Staubli VAL3: valGI.pjx

--- valGI.pjx ---
Parameters version=s8.15.3Cs9_BS3337 stackSize=200000 millimeterUnit=true
Program file=_getForce.pgx
Program file=_productCycle.pgx
Program file=_tCycleCtrl.pgx
Program file=createUserTask.pgx
Program file=cycle_Abort.pgx
Program file=cycle_End.pgx
Program file=cycle_GoHome.pgx
Program file=cycle_Hold.pgx
Program file=cycle_Init.pgx
Program file=cycle_Reset.pgx
Program file=cycle_RotGoHome.pgx
Program file=cycle_Start.pgx
Program file=cycle_Stop.pgx
Program file=cycle_Unhold.pgx
Program file=Init.pgx
Program file=kill.pgx
Program file=Main.pgx
Program file=MonitorIO.pgx
Program file=MonitorIO1.pgx
Program file=start.pgx
Program file=stop.pgx
Data file=valGI.dtx
Library alias=rs path=Disk://source/projectSource/robotStatus/robotStatus.pjx
Library alias=io path=Disk://source/projectSource/io/io.pjx
Library alias=act path=Disk://source/projectSource/Action/Action.pjx
Library alias=savedata path=Disk://source/saveData/saveData.pjx
Library alias=home path=Disk://HMI_cs9/home/home.pjx
Library alias=plc path=Disk://source/projectSource/plc/plc.pjx
Library alias=prog path=Disk://source/projectSource/program/program.pjx
Library alias=safeHome path=Disk://source/projectSource/goSafeHome/goSafeHome.pjx
Library alias=safe path=Disk://safeLogic/safeLogic.pjx
Library alias=program path=Disk://source/projectSource/program/program.pjx
Library alias=hmi_util path=Disk://HMI_cs9/HMI_util/HMI_util.pjx
Library alias=saveData path=Disk://source/saveData/saveData.pjx
Library alias=initLib path=./initLib/initLib.pjx
Library alias=libTqe path=Disk://LibTorque/LibTorque.pjx
Library alias=trajectory path=Disk://source/projectSource/trajectory/trajectory.pjx
Library alias=ar path=Disk://autoReturn/autoReturn.pjx

--- valGI.dtx ---
bool _bAtHome
bool _bEndCycle
bool _bHeavyAlarm
bool _bIsScara
bool _bShowEndBt
bool _bShowPauseBt
bool _bShowResetBt
bool _bShowStartBt
bool _bShowStopBt
bool bBool
bool bControlByRobot = true
bool bTosave
frame test3 = {fatherId=world[0]}
num _nAvgCapacity
num _nBestCapacity
num _nCTIndex
num _nCapacity
num _nClock[10]
  [1] = 12488.271809
  [3] = 12488.271821
num _nCycleTime[10]
num _nLastStateCMD
num _nOmacStat
num _nStateCMD
num nCycleCmd
num nErrorCode = 1
num nLastLib
num nProgCode
string _sArmType
string _sOmacCmd
string _sOmacStatus = "1"
string _sPageAvergeCapacity
string _sPageBestCapacity
string _sPageCurrentCapacity
string _sPageCycleStatus
string _sPageHerej
string _sPagePosition
string _sPageProfile
string _sPageRobotStatus
string _sPageSN
string sMsg
num nForce[6]
public bool bGetMovId
mdesc mHome = {accel=20, vel=20, decel=20, blend=off}

--- Main.pgx ---
program Main()
  local bool l_bResult
  local bool l_bStartClock
  local num l_nClock
  local num l_nResult
begin
  //

  home:sVersion="version:4.11.20251028"
  resetMotion()
  //初始化
  call cycle_Init()


  //
  userPage("StartUp")

  sMsg=">>> Loading 数据库 "+toString("",savedata:nLibIndex)+" <<<"
  //guohangxin add 2023.03.23
  call initLib:initlib()
  call program:loadPROG(saveData:nLibIndex,l_nResult)
  call trajectory:loadTRAJ(saveData:nLibIndex,l_nResult)
  sMsg=""
  //机器人控制任务
  taskCreate "cycleCtrl",90,_tCycleCtrl()
  wait(taskStatus("cycleCtrl")==1)
  //机器人状态
  taskCreate "plc",60,plc:main()
  wait(taskStatus("plc")==1)
  //HMI
  taskCreate "HMI",50,home:main()
  wait(taskStatus("HMI")==1)
  //lifebit
  taskCreate "lifebit",10,plc:lifebit()
  wait(taskStatus("lifebit")==1)
  //创建用户自定义的任务
  //call createUserTask()
  //safe check
  taskCreate "safeCheck",80,safe:main()
  wait(taskStatus("safeCheck")==1)
  do
    //任务监控
    if taskStatus("plc")>1 and (clock()-_nClock[1]>5)
      _nClock[1]=clock()
      taskResume("plc",1)
    else
      _nClock[1]=clock()
    endIf
    if taskStatus("HMI")>1
      //保存当前数据
      bTosave=true
      call trajectory:onSave(bTosave)
      bTosave=true
      call program:onSave(bTosave)
      wait(rs:bIsSaving==false)
      l_bResult=userPageConfirm("需要重载HMI应用？")
      if l_bResult

        taskKill("HMI")
        wait(taskStatus("HMI")==-1)
        taskCreate "HMI",50,home:main()
        wait(taskStatus("HMI")==1)
      endIf
    endIf
    if taskStatus("lifebit")>1 and (clock()-_nClock[3]>5)
      _nClock[3]=clock()
      taskResume("lifebit",1)
    else
      _nClock[3]=clock()
    endIf

    delay(0)
  until rs:bQuitApp==true

  call kill()

end

--- start.pgx ---
program start()
begin
  taskCreate "appMain",20,Main()
end

--- _getForce.pgx ---
program _getForce()
  local num i
  local num l_nForce[6]
begin
  for i=0 to 5
    nForce[i]=0
  endFor

  do
    getJointForce(l_nForce)
    for i=0 to 5
      if abs(l_nForce[i])>nForce[i]
        nForce[i]=abs(l_nForce[i])
      endIf
    endFor
    //      if abs(l_nForce[4])>nForce[4]
    //        nForce[4]=abs(l_nForce[4])
    //      endIf
    //      if abs(l_nForce[5])>nForce[5]
    //        nForce[5]=abs(l_nForce[5])
    //      endIf
    delay(0)
  until rs:_nOmacStat==1
  //logMsg("程序号"+toString(".",rs:nProgCode)+"最大J5扭矩："+toString(".3",nForce[4])+",最大J6扭矩："+toString(".3",nForce[5]))
  rs:_sRobotStatus="程序号:"+toString(".",rs:nProgCode)+",J1MaxForce："+toString(".2",nForce[0])+",J2MaxForce："+toString(".2",nForce[1])+",J3MaxForce："+toString(".2",nForce[2])+",J4MaxForce："+toString(".2",nForce[3])+",J5MaxForce："+toString(".2",nForce[4])+",J6MaxForce："+toString(".2",nForce[5])
end

--- _productCycle.pgx ---
public program _productCycle()
  local bool l_bErr
  local bool l_bStartClock
  local num l_nClock
  local num l_nLastAct
  local num l_nLibIndex
  local string l_sPath
begin
  //do
  // rs:nPLCcmd=0
  //等待数据库切换完成以及程序号完成
  // wait(io:dInput[30]==true)
  //wait(bBool==true)
  //
  waitEndMove()
  //
  //（工作号&程序号->切换完成->plc启动信号->productcycle->（工作号&程序号->切换完成->plc启动信号
  //
  //获取程序号
  call io:getAnaIO(io:aInItem[0].aAio,rs:nProgCode,l_bErr)
  switch rs:nProgCode
    case 0
      //call prog:makeTraj("test")
    break
    case 1
      rs:sTrajStatus="开始执行prod01"
      call prog:makeTraj("prod01")

    break
    case 2
      rs:sTrajStatus="开始执行prod02"
      call prog:makeTraj("prod02")

    break
    case 3
      rs:sTrajStatus="开始执行prod03"
      call prog:makeTraj("prod03")

    break
    case 4
      rs:sTrajStatus="开始执行prod04"
      call prog:makeTraj("prod04")

    break
    case 5
      rs:sTrajStatus="开始执行prod05"
      call prog:makeTraj("prod05")

    break
    case 6
      rs:sTrajStatus="开始执行prod06"
      call prog:makeTraj("prod06")

    break
    case 7
      rs:sTrajStatus="开始执行prod07"
      call prog:makeTraj("prod07")

    break
    case 8
      rs:sTrajStatus="开始执行prod08"
      call prog:makeTraj("prod08")

    break
    case 9
      rs:sTrajStatus="开始执行prod09"
      call prog:makeTraj("prod09")

    break
    case 10
      rs:sTrajStatus="开始执行prod10"
      call prog:makeTraj("prod10")

    break
    case 11
      rs:sTrajStatus="开始执行prod11"
      call prog:makeTraj("prod11")

    break
    case 12
      rs:sTrajStatus="开始执行prod012"
      call prog:makeTraj("prod12")

    break
    case 13
      rs:sTrajStatus="开始执行prod13"
      call prog:makeTraj("prod13")

    break
    case 14
      rs:sTrajStatus="开始执行prod14"
      call prog:makeTraj("prod14")

    break
    case 15
      rs:sTrajStatus="开始执行prod15"
      call prog:makeTraj("prod15")

    break
    case 16
      rs:sTrajStatus="开始执行prod16"
      call prog:makeTraj("prod16")

    break


    case 17
      rs:sTrajStatus="开始执行prod17"
      call prog:makeTraj("prod17")
    break

    case 18
      rs:sTrajStatus="开始执行prod18"
      call prog:makeTraj("prod18")
    break
    case 19
      rs:sTrajStatus="开始执行prod19"
      call prog:makeTraj("prod19")
    break

    case 20
      rs:sTrajStatus="开始执行prod20"
      call prog:makeTraj("prod20")
    break

    case 21
      rs:sTrajStatus="开始执行prod21"
      call prog:makeTraj("prod21")

    break
    case 22
      rs:sTrajStatus="开始执行prod22"
      call prog:makeTraj("prod22")

    break
    case 23
      rs:sTrajStatus="开始执行prod23"
      call prog:makeTraj("prod23")

    break
    case 24
      rs:sTrajStatus="开始执行prod24"
      call prog:makeTraj("prod24")

    break
    case 25
      rs:sTrajStatus="开始执行prod25"
      call prog:makeTraj("prod25")

    break
    case 26
      rs:sTrajStatus="开始执行prod26"
      call prog:makeTraj("prod26")

    break
    case 27
      rs:sTrajStatus="开始执行prod27"
      call prog:makeTraj("prod27")

    break
    case 28
      rs:sTrajStatus="开始执行prod28"
      call prog:makeTraj("prod28")

    break
    case 29
      rs:sTrajStatus="开始执行prod29"
      call prog:makeTraj("prod29")

    break
    case 30
      rs:sTrajStatus="开始执行prod30"
      call prog:makeTraj("prod30")

    break
    case 31
      rs:sTrajStatus="开始执行prod31"
      call prog:makeTraj("prod31")

    break
    case 32
      rs:sTrajStatus="开始执行prod032"
      call prog:makeTraj("prod32")

    break
    case 33
      rs:sTrajStatus="开始执行prod33"
      call prog:makeTraj("prod33")

    break
    case 34
      rs:sTrajStatus="开始执行prod34"
      call prog:makeTraj("prod34")

    break
    case 35
      rs:sTrajStatus="开始执行prod35"
      call prog:makeTraj("prod35")

    break
    case 36
      rs:sTrajStatus="开始执行prod36"
      call prog:makeTraj("prod36")

    break

    case 37
      rs:sTrajStatus="开始执行prod37"
      call prog:makeTraj("prod37")
    break

    case 38
      rs:sTrajStatus="开始执行prod38"
      call prog:makeTraj("prod38")
    break
    case 39
      rs:sTrajStatus="开始执行prod39"
      call prog:makeTraj("prod39")
    break

    case 40
      rs:sTrajStatus="开始执行prod40"
      call prog:makeTraj("prod40")
    break
    case 40
      rs:sTrajStatus="开始执行prod40"
      call prog:makeTraj("prod40")

    break
    case 41
      rs:sTrajStatus="开始执行prod41"
      call prog:makeTraj("prod41")

    break
    case 42
      rs:sTrajStatus="开始执行prod042"
      call prog:makeTraj("prod42")

    break
    case 43
      rs:sTrajStatus="开始执行prod43"
      call prog:makeTraj("prod43")

    break
    case 44
      rs:sTrajStatus="开始执行prod44"
      call prog:makeTraj("prod44")

    break
    case 45
      rs:sTrajStatus="开始执行prod45"
      call prog:makeTraj("prod45")

    break
    case 46
      rs:sTrajStatus="开始执行prod46"
      call prog:makeTraj("prod46")

    break

    case 47
      rs:sTrajStatus="开始执行prod47"
      call prog:makeTraj("prod47")
    break

    case 48
      rs:sTrajStatus="开始执行prod48"
      call prog:makeTraj("prod48")
    break
    case 49
      rs:sTrajStatus="开始执行prod49"
      call prog:makeTraj("prod49")
    break

    case 50
      rs:sTrajStatus="开始执行prod50"
      call prog:makeTraj("prod50")
    break

  endSwitch
  if l_bStartClock and l_nLastAct!=rs:nActCode
    rs:_nCTIndex=(rs:_nCTIndex+1)%size(rs:_nCycleTime)
    rs:_nCycleTime[rs:_nCTIndex]=clock()-l_nClock
  else
    l_bStartClock=true
  endIf
  l_nClock=clock()
  l_nLastAct=rs:nActCode
  //delay(0)
  //
  rs:_nOmacStat=1
  rs:sTrajStatus=""
  rs:_sRobotStatus="当前件生产结束"
  //2025.1.6 add 结束扭矩记录程序
  if taskStatus("getForce")!=-1
    delay(0.2)
    taskKill("getForce")
  endIf
end

--- _tCycleCtrl.pgx ---
program _tCycleCtrl()
  local bool l_bAckAlarm
  local bool l_bEndCmd
  local bool l_bErr
  local bool l_bHoldCmd
  local bool l_bPowerOff
  local bool l_bPowerOn
  local bool l_bResetCmd
  local bool l_bResetIO
  local bool l_bStartCmd
  local bool l_bStopCmd
  local num l_n
begin
  //  rs:_nOmacStat
  //1-Ready
  //2-Starting
  //3-Running
  //4-Resetting
  //5-Holding
  //6-Held
  //7-Ending
  //8-Stopping
  //9-Stopped
  //10-Aborting

  // _nStateCmd
  //1-Reset
  //2-Start
  //3-Hold
  //4-Unhold
  //5-End
  //6-Stop
  //7-Abort

  do
    //add by guohangxin 20240408 refreshing log
    call rs:robotStatus()
    //    if rs:bIsHome and workingMode()==4 and esStatus()!=2 and rs:_nOmacStat==9
    //      rs:_nOmacStat=1
    //    endIf
    //****************************Cycle control*****************************//
    //7-Abort
    if rs:_bHeavyAlarm==true and (rs:_nOmacStat<9 and rs:_nOmacStat!=3 and rs:_nOmacStat!=6) or (workingMode()==1 and rs:_nOmacStat<9)
      //********add by guohangxin log**********//
      if rs:_bHeavyAlarm==true
        rs:_sRobotStatus="当前机器人有报警,代码:"+toString("",rs:_nAlarmCode[rs:_nErrIndex])
      elseIf(workingMode()==1 and rs:_nOmacStat<9)
        rs:_sRobotStatus="当前机器人处于手动非停止状态"
      endIf
      //***************************************//
      _nStateCMD=7
      //1-Reset
    elseIf(rs:nPLCcmd==1 or rs:nCycleCmd==1) and rs:_nOmacStat==9
      //********add by guohangxin log**********//
      if rs:nPLCcmd==1
        rs:_sRobotStatus="收到PLC复位信号"
      elseIf rs:nCycleCmd==1
        rs:_sRobotStatus="页面设置复位信号"
      endIf
      if rs:_bHeavyAlarm==false
        _nStateCMD=1
      else
        _nStateCMD=0
        popUpMsg("请先清除报错!")
        delay(3)
      endIf
      //***************************************//
      //2-Start
    elseIf(rs:nPLCcmd==2 or rs:nCycleCmd==2) and rs:_nOmacStat==1
      //********add by guohangxin log**********//
      if rs:nPLCcmd==2
        rs:_sRobotStatus="收到PLC启动信号"
      elseIf rs:nCycleCmd==2
        rs:_sRobotStatus="页面设置启动信号"
      endIf
      if rs:_bHeavyAlarm==false
        _nStateCMD=2
      else
        _nStateCMD=0
        popUpMsg("请先清除报错!")
        delay(3)
      endIf
      //***************************************//
      //3-Hold
    elseIf(rs:nPLCcmd==3 or rs:nCycleCmd==3 or rs:_bHeavyAlarm==true) and rs:_nOmacStat==3
      //********add by guohangxin log**********//
      if rs:nPLCcmd==3
        rs:_sRobotStatus="收到PLC暂停信号"
      elseIf rs:nCycleCmd==3
        rs:_sRobotStatus="页面设置暂停信号"
      elseIf rs:_bHeavyAlarm==true
        rs:_sRobotStatus="机器人报警，暂停生产"
      endIf
      //***************************************//
      _nStateCMD=3
      //4-Unhold
    elseIf(rs:nPLCcmd==2 or rs:nCycleCmd==4) and rs:_nOmacStat==6
      //********add by guohangxin log**********//
      if rs:nPLCcmd==2
        rs:_sRobotStatus="收到PLC暂停恢复信号"
      elseIf rs:nCycleCmd==4
        rs:_sRobotStatus="页面设置暂停恢复信号"
      endIf
      //***************************************//
      if rs:_bHeavyAlarm==false
        _nStateCMD=4
      else
        _nStateCMD=0
        popUpMsg("请先清除报错!")
        delay(3)
      endIf
      //5-End
    elseIf(rs:nPLCcmd==4 or rs:nCycleCmd==5) and rs:_nOmacStat==3
      //********add by guohangxin log**********//
      if rs:nPLCcmd==4
        rs:_sRobotStatus="收到PLC生产结束信号"
      elseIf rs:nCycleCmd==5
        rs:_sRobotStatus="页面设置生产结束信号"
      endIf
      //***************************************//
      _nStateCMD=5
      //6-Stop
    elseIf(rs:nPLCcmd==5 or rs:nCycleCmd==6) and rs:_nOmacStat<8
      //********add by guohangxin log**********//
      if rs:nPLCcmd==5
        rs:_sRobotStatus="收到PLC停止信号"
      elseIf rs:nCycleCmd==6
        rs:_sRobotStatus="页面设置停止信号"
      endIf
      //***************************************//
      _nStateCMD=6
      //2025.7.21 add 增加路径回原程序
      //elseIf(rs:nPLCcmd==6) and (rs:_nOmacStat==9 and rs:_nOmacStat!=11) and rs:bIsHome==false and esStatus()!=2 and workingMode()==4
    elseIf (rs:nCycleCmd==7 or rs:nPLCcmd==7) and (rs:_nOmacStat==9 and rs:_nOmacStat!=11) and rs:bIsHome==false and esStatus()!=2 and (workingMode()==4 or workingMode()==1)
      if rs:_bHeavyAlarm==false and ioStatus(io:dORbHeartbeat)>=0
        if rs:nPLCcmd==7
          rs:_sRobotStatus="收到PLC路径回Home点信号"
        elseIf rs:nCycleCmd==7
          rs:_sRobotStatus="收到页面手动路径回Home点信号"
        endIf
        _nStateCMD=8
      else
        _nStateCMD=0
        popUpMsg("请先清除报错!")
        delay(3)
      endIf
      //2025.7.21 add 增加直接回原程序
    elseIf (rs:nPLCcmd==6) and ((rs:_nOmacStat==9 or rs:_nOmacStat==11) and rs:_nOmacStat!=12) and rs:bIsHome==false and esStatus()!=2 and workingMode()==4
      if rs:_bHeavyAlarm==false and ioStatus(io:dORbHeartbeat)>=0
        rs:_sRobotStatus="收到PLC直接回Home点信号"
        _nStateCMD=9
      else
        _nStateCMD=0
        popUpMsg("请先清除报错!")
        delay(3)
      endIf
    else
      _nStateCMD=0
    endIf

    //if _nStateCMD!=_nLastStateCMD
    switch _nStateCMD
      //Reset
      case 1
        if rs:_nOmacStat==9
          if taskStatus("Reset")>=0
            taskKill("Reset")
          endIf
          wait(taskStatus("Reset")<0)
          delay(0.1)
          taskCreate "Reset",100,cycle_Reset()
        endIf
      break

      //Start
      case 2
        if rs:_nOmacStat==1
          if taskStatus("Start")>=0
            taskKill("Start")
          endIf
          wait(taskStatus("Start")<0)
          delay(0.1)
          taskCreate "Start",100,cycle_Start()
        endIf
      break

      //Hold
      case 3
        if taskStatus("Hold")>=0
          taskKill("Hold")
        endIf
        wait(taskStatus("Hold")<0)
        taskCreate "Hold",100,cycle_Hold()
      break

      //unHold
      case 4
        if taskStatus("Unhold")>=0
          taskKill("Unhold")
        endIf
        wait(taskStatus("Unhold")<0)
        taskCreate "Unhold",100,cycle_Unhold()
        delay(0.1)
      break

      case 5
        if taskStatus("End")>=0
          taskKill("End")
        endIf
        wait(taskStatus("End")<0)
        taskCreate "End",100,cycle_End()
      break

      //Stop
      case 6
        if taskStatus("Stop")>=0
          taskKill("Stop")
        endIf
        wait(taskStatus("Stop")<0)
        taskCreate "Stop",100,cycle_Stop()
      break

      //Abort
      case 7
        if taskStatus("Abort")>=0
          taskKill("Abort")
        endIf
        wait(taskStatus("Abort")<0)
        taskCreate "Abort",100,cycle_Abort()
      break
            //路径回Home
      case 8
        if taskStatus("RotGoHome")>=0
          taskKill("RotGoHome")
        endIf
        wait(taskStatus("RotGoHome")<0)
        taskCreate "RotGoHome",100,cycle_RotGoHome()
      break

      //直接回Home
      case 9
        if taskStatus("GoHome")>=0
          taskKill("GoHome")
        endIf
        wait(taskStatus("GoHome")<0)
        taskCreate "GoHome",100,cycle_GoHome()
      break
    endSwitch
    // endIf
    //记录上次指令
    //_nLastStateCMD=_nStateCMD
    delay(0.02)
  until false
end

--- createUserTask.pgx ---
program createUserTask()
begin
  //作用：调用自定义的任务
  //1.创建动作Action任务
  call act:create()
  //2.创建视觉任务
end

--- cycle_Abort.pgx ---
program cycle_Abort()
begin
  // abort task
  rs:_nOmacStat=10
  taskKill("GoHome")
  taskKill("Monitor")
  taskKill("RotGoHome")
  taskKill("Monitor1")
  call ar:getCurMoveID(bGetMovId,"Abort")
  stopMove()
  resetMotion()

  // Stop task
  taskKill("Reset")
  taskKill("Start")
  taskKill("Stop")
  taskKill("End")
  taskKill("productCycle")
  taskKill("getForce")
  wait(isSettled())
  disablePower()
  wait(isPowered()==false)
    //2025.7.21 add 复位输出信号
  call plc:resetOutput()
  //OMAC进程:Stopped
  rs:_nOmacStat=9
  logMsg("当前处于生产停止状态 "+toString(".2",clock()))
  rs:_sRobotStatus="当前处于生产停止状态"
  delay(0)
end

--- cycle_End.pgx ---
program cycle_End()
begin

  //cycle进程:Ending
  rs:_nOmacStat=7
  _bEndCycle=true
  wait(taskStatus("Main")<0)

  // Stop task
  stopMove()
  call ar:getCurMoveID(bGetMovId,"End")
  wait(isSettled())
  resetMotion()
  //shutdown arm power
  disablePower()

  //cycle进程:Stopped
  rs:_nOmacStat=9
  logMsg("当前处于停止状态 "+toString(".2",clock()))
  rs:_sRobotStatus="当前处于停止状态"
end

--- cycle_GoHome.pgx ---
program cycle_GoHome()
  local tool l_tTool
begin
  rs:_nOmacStat=12
  // Stop task
  taskKill("Reset")
  taskKill("Start")
  taskKill("Stop")
  taskKill("End")
  taskKill("Monitor1")
  taskKill("RotGoHome")
  taskKill("productCycle")

  wait(isSettled())

  if !isPowered()
    popUpMsg("请先上电！")
    rs:_nOmacStat=9
    return
  endIf

  resetMotion()
  //2024.11.22 add初始化回零堆栈
  call ar:resetReturnStack(false)
  rs:sTrajStatus="直接回原点过程中"
  taskCreate "Monitor",20,MonitorIO()
  wait(taskStatus("Monitor")==1)
  link(l_tTool,flange)
  call saveData:getTool(1,l_tTool)
  movej(saveData:jHome,l_tTool,mHome)
  waitEndMove()
  ar:bInterrupt=false
  bGetMovId=false
  rs:sTrajStatus="直接回原点完成"

  taskKill("Monitor")
  wait(taskStatus("Monitor")<0)
  disablePower()
  rs:_nOmacStat=9
  delay(0)

end

--- cycle_Hold.pgx ---
program cycle_Hold()
begin
  //cycle进程:Holding
  rs:_nOmacStat=5
  //if isPowered()
  //    disablePower()
  //    watch(isPowered()==false,2)
  //  endIf
  stopMove()
  wait(isSettled())
  //cycle进程:Held
  rs:_nOmacStat=6
  logMsg("当前处于暂停状态 "+toString(".2",clock()))
  rs:_sRobotStatus="当前处于暂停状态"
end

--- cycle_Init.pgx ---
program cycle_Init()
begin
  //
  call Init()
  //
  call act:init()
  //
  call io:init()

  //  if !isPowered() and workingMode()==4
  //    enablePower()
  //    delay(1)
  //  endIf

end

--- cycle_Reset.pgx ---
program cycle_Reset()
  local bool l_bEdge
begin
  setSafetyRestart()
  delay(0.1)
  //进程:resetting
  rs:_nOmacStat=4

  taskKill("Start")
  taskKill("Stop")
  taskKill("End")
  taskKill("Main")
  taskKill("GoHome")
  taskKill("Monitor")
  taskKill("RotGoHome")
  taskKill("Monitor1")


  call rs:init()
  call ar:getCurMoveID(bGetMovId,"Reset")
  resetMotion()

  // Enables arm power
  do
    if workingMode()==4
      enablePower()
      delay(1)
    elseIf workingMode()==1 and l_bEdge==false
      l_bEdge=true
      popUpMsg("当前工作模式为手动，请手动上电")
    endIf
  until isPowered()==true
  //2025.1.6 add 设置扭矩保护
  call libTqe:_setMaxJntForce()
  if !rs:bIsHome
    popUpMsg("请手动回原点")
    return
  endIf
  //回home
  //call safeHome:gosafe()
  prog:nLastIndex=0

  //进程:ready
  rs:_nOmacStat=1
  logMsg("当前处于ready状态 "+toString(".2",clock()))
  rs:_sRobotStatus="当前处于ready状态"
  delay(0)
end

--- cycle_RotGoHome.pgx ---
program cycle_RotGoHome()
  local bool l_bContain
begin
  //  stopMove()
  //  resetMotion()
  //检查堆栈是否存有点位
  call ar:getMotCount(l_bContain)
  if !l_bContain
    //popUpMsg("无法路径回原，请手动回原点！")
    return
  endIf

  rs:_nOmacStat=11
  // Stop task
  taskKill("Reset")
  taskKill("Start")
  taskKill("Stop")
  taskKill("End")
  taskKill("GoHome")
  taskKill("Monitor")
  taskKill("productCycle")

  wait(isSettled())
  //  if !isPowered()
  //    enablePower()
  //    wait(isPowered()==true)
  //  endIf
  if !isPowered()
    popUpMsg("请先手动上电！")
    rs:_nOmacStat=9
    return
  endIf

  //2024.12.02 add 监控IO程序
  rs:sTrajStatus="路径回原点过程中"
  if rs:nCycleCmd!=7
    taskCreate "Monitor1",20,MonitorIO1()
    wait(taskStatus("Monitor1")==1)
  endIf

  call ar:returnMove(false,savedata:jHome,bGetMovId)


  if rs:bIsHome
    rs:sTrajStatus="路径回原点完成"
    bGetMovId=false
    ar:bInterrupt=false
  endIf

  if rs:nCycleCmd!=7
    taskKill("Monitor1")
    wait(taskStatus("Monitor1")<0)
  endIf
  disablePower()
  rs:_nOmacStat=9
  delay(0)

end

--- cycle_Start.pgx ---
program cycle_Start()
  local bool l_bErr
begin

  //OMAC进程:Starting
  rs:_nOmacStat=2
  //运行startUp程序
  waitEndMove()
  call io:getAnaIO(io:aInItem[0].aAio,rs:nProgCode,l_bErr)

  //切换数据库
  //  savedata:nLibIndex=aioGet(io:aInput[2])
  //  delay(0)
  //  call plc:changeDataLib1(savedata:nLibIndex)
  //  aioSet(io:aOutput[3],savedata:nLibIndex)

  //2025.1.6 add 开始扭矩记录程序，获取实时扭矩
  if taskStatus("getForce")>=0
    taskKill("getForce")
    wait(taskStatus("getForce")<0)
  endIf
  taskCreate "getForce",100,_getForce()
  wait(taskStatus("getForce")==1)
  //创建生产任务
  if taskStatus("productCycle")>=0
    taskKill("productCycle")
    wait(taskStatus("productCycle")<0)
  endIf
  taskCreate "productCycle",100,_productCycle()
  wait(taskStatus("productCycle")==1)
  //OMAC进程:Start
  rs:_nOmacStat=3
  logMsg("当前处于生产状态 "+toString(".2",clock()))
  rs:_sRobotStatus="当前处于生产状态"
end

--- cycle_Stop.pgx ---
program cycle_Stop()
begin
  //进程:Stopping
  rs:_nOmacStat=8
  // Stop task
  taskKill("Reset")
  taskKill("Start")
  taskKill("productCycle")
  taskKill("End")
  taskKill("GoHome")
  taskKill("Monitor")
  taskKill("RotGoHome")
  taskKill("Monitor1")
  taskKill("getForce")

  while !isPowered()
    enablePower()
    delay(1)
  endWhile
  //
  stopMove()
  call ar:getCurMoveID(bGetMovId,"Stop")
  resetMotion()
  disablePower()
  wait(isPowered()==false)
  //2025.7.21 add 复位输出信号
  call plc:resetOutput()
  //OMAC进程:Stopped
  rs:_nOmacStat=9
  logMsg("当前处于生产停止状态 "+toString(".2",clock()))
  rs:_sRobotStatus="当前处于生产停止状态"
  delay(0)
end

--- cycle_Unhold.pgx ---
program cycle_Unhold()
begin
  //cycle进程:unholding
  rs:_nOmacStat=2
  //enable power
  if !isPowered()
    enablePower()
    watch(isPowered(),2)
  endIf
  restartMove()
  //cycle进程:running
  rs:_nOmacStat=3
  logMsg("当前处于生产状态 "+toString(".2",clock()))
  rs:_sRobotStatus="当前处于生产状态"
end

--- Init.pgx ---
program Init()
  local num i
  local string l_sArmType
begin
  //dio

  //****************bool*****************
  _bEndCycle=false
  _bAtHome=false
  _bHeavyAlarm=false
  //判断是否是4轴机器人
  l_sArmType=left(getVersion("Arm Type"),2)
  _bIsScara=(l_sArmType=="rs" or l_sArmType=="ts" or l_sArmType=="tp")


  call rs:init()

end

--- kill.pgx ---
program kill()
begin
  //kill all task
  taskKill("safeCheck")
  taskKill("Reset")
  taskKill("Start")
  taskKill("Stop")
  taskKill("cycleCtrl")
  taskKill("plc")
  taskKill("lifebit")
  taskKill("actCtrl")
  taskKill("appMain")
  taskKill("HMI")

  //
  rs:bQuitApp=false
  stopMove()
  resetMotion()
  disablePower()
end

--- MonitorIO.pgx ---
program MonitorIO()
  local bool l_bStopMove
  local bool l_bToHome
  local bool l_bRestartMove
  local bool l_bErr
begin
  l_bRestartMove=true
  l_bStopMove=false
  do
    call io:getDigIO(io:dInput[9],l_bToHome,l_bErr)
    if l_bToHome and (!l_bRestartMove or l_bStopMove)
      l_bRestartMove=true
      l_bStopMove=false
      restartMove()
    endIf

    if !l_bToHome and !l_bStopMove
      l_bStopMove=true
      stopMove()
    endIf

//    if manual:bJogMove
//      if taskStatus("GoHome")>=0
//        taskKill("GoHome")
//      endIf
//      wait(taskStatus("GoHome")<0)

//      stopMove()
//      resetMotion()
//      rs:_nOmacStat=9
//      taskKill("Monitor")
//      wait(taskStatus("Monitor")<0)
//    endIf
    delay(0)
  until false

end

--- MonitorIO1.pgx ---
program MonitorIO1()
  local bool l_bStopMove
  local bool l_bToHome
  local bool l_bRestartMove
  local bool l_bErr
begin
  l_bRestartMove=true
  l_bStopMove=false
  do
    call io:getDigIO(io:dInput[10],l_bToHome,l_bErr)
    if l_bToHome and (!l_bRestartMove or l_bStopMove)
      l_bRestartMove=true
      l_bStopMove=false
      restartMove()
    endIf

    if !l_bToHome and !l_bStopMove
      l_bStopMove=true
      stopMove()
    endIf

//    if manual:bJogMove
//      if taskStatus("RotGoHome")>=0
//        taskKill("RotGoHome")
//      endIf
//      wait(taskStatus("RotGoHome")<0)

//      stopMove()
//      resetMotion()
//      //2024.11.22 add初始化回零堆栈
//      call ar:resetReturnStack(false)
//      rs:_nOmacStat=9
//      taskKill("Monitor1")
//      wait(taskStatus("Monitor1")<0)
//    endIf
    delay(0)
  until false

end

--- stop.pgx ---
program stop()
begin
  //kill all task
  taskKill("Reset")
  taskKill("Start")
  taskKill("Stop")
  taskKill("cycleCtrl")
  taskKill("Zones")
  taskKill("Main")
  taskKill("StatusRobot")
  //
  stopMove()
  resetMotion()
  disablePower()
end
